(* CODESYS project ManualRequest.xml

Project tree, tasks and I/O mapping:
  visualisation ManualRequest
*)

// /ManualRequest
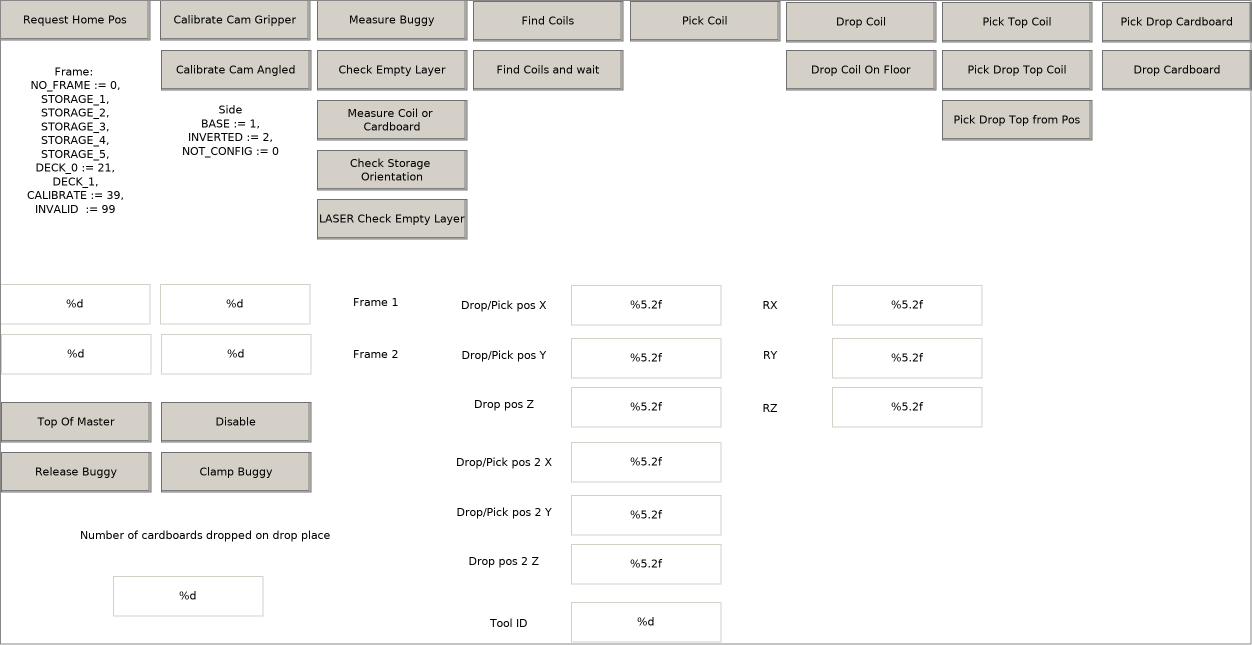
VISUALIZATION ManualRequest  // 1252x645
    Button (160,0 150x40), "Calibrate Cam Gripper", input disabled if: NOT PRG_VisuTask_10ms._fbManualCtrl.xManualMode
        tap PRG_VisuTask_10ms._fbManualCtrl._btnCalibrateCamGripper.xbtn
    Button (0,0 150x40), "Request Home Pos", input disabled if: NOT PRG_VisuTask_10ms._fbManualCtrl.xManualMode
        tap PRG_VisuTask_10ms._fbManualCtrl._btnRequestHomePos.xbtn
    Button (317,0 150x40), "Measure Buggy", input disabled if: NOT PRG_VisuTask_10ms._fbManualCtrl.xManualMode
        tap PRG_VisuTask_10ms._fbManualCtrl._btnMeasure.xbtn
    Textfield (0,284 150x40), "%d", text variable: PRG_VisuTask_10ms._fbManualCtrl._scRobotPosition.eStorage
        OnMouseUp: write the text variable via Default
    Textfield (160,284 150x40), "%d", text variable: PRG_VisuTask_10ms._fbManualCtrl._scRobotPosition.eSide
        OnMouseUp: write the text variable via Default
    Label (0,50 151x181), "Frame: NO_FRAME := 0, STORAGE_1, STORAGE_2, STORAGE_3, STORAGE_4, STORAGE_5, DECK_0 := 21, DECK_1, CALIBRATE := 39, INVALID := 99"
    Label (160,50 141x161), "Side BASE := 1, INVERTED := 2, NOT_CONFIG := 0"
    Button (473,1 150x40), "Find Coils", input disabled if: NOT PRG_VisuTask_10ms._fbManualCtrl.xManualMode
        tap PRG_VisuTask_10ms._fbManualCtrl._btnFindCoils.xbtn
    Button (630,1 150x40), "Pick Coil", input disabled if: NOT PRG_VisuTask_10ms._fbManualCtrl.xManualMode
        tap PRG_VisuTask_10ms._fbManualCtrl._btnPickCoil.xbtn
    Button (1,402 150x40), "Top Of Master", input disabled if: NOT PRG_VisuTask_10ms._fbManualCtrl.xManualMode
        tap PRG_VisuTask_10ms._fbManualCtrl._btnRequestTopOfMaster.xbtn
    Button (161,402 150x40), "Disable", input disabled if: NOT PRG_VisuTask_10ms._fbManualCtrl.xManualMode
        tap PRG_VisuTask_10ms._fbManualCtrl._btnRequestDisable.xbtn
    Button (786,2 150x40), "Drop Coil", input disabled if: NOT PRG_VisuTask_10ms._fbManualCtrl.xManualMode
        tap PRG_VisuTask_10ms._fbManualCtrl._btnDropCoil.xbtn
    Button (942,2 150x40), "Pick Top Coil", input disabled if: NOT PRG_VisuTask_10ms._fbManualCtrl.xManualMode
        tap PRG_VisuTask_10ms._fbManualCtrl._btnPickTopCoil.xbtn
    Button (1,452 150x40), "Release Buggy", input disabled if: NOT PRG_VisuTask_10ms._fbManualCtrl.xManualMode
        tap PRG_VisuTask_10ms._fbManualCtrl._btnReleaseBuggy.xbtn
    Button (161,452 150x40), "Clamp Buggy", input disabled if: NOT PRG_VisuTask_10ms._fbManualCtrl.xManualMode
        tap PRG_VisuTask_10ms._fbManualCtrl._btnClampBuggy.xbtn
    Label (445,284 118x43), "Drop/Pick pos X"
    Textfield (571,285 150x40), "%5.2f", text variable: PRG_VisuTask_10ms._fbManualCtrl._scRobotPosition.scRobotPosition.posX
        OnMouseUp: write the text variable via Default
    Textfield (571,338 150x40), "%5.2f", text variable: PRG_VisuTask_10ms._fbManualCtrl._scRobotPosition.scRobotPosition.posY
        OnMouseUp: write the text variable via Default
    Label (445,334 118x43), "Drop/Pick pos Y"
    Label (445,383 118x43), "Drop pos Z"
    Textfield (571,387 150x40), "%5.2f", text variable: PRG_VisuTask_10ms._fbManualCtrl._scRobotPosition.scRobotPosition.posZ
        OnMouseUp: write the text variable via Default
    Button (786,50 150x40), "Drop Coil On Floor", input disabled if: NOT PRG_VisuTask_10ms._fbManualCtrl.xManualMode
        tap PRG_VisuTask_10ms._fbManualCtrl._btnDropCoilOnFloor.xbtn
    Button (942,50 150x40), "Pick Drop Top Coil", input disabled if: NOT PRG_VisuTask_10ms._fbManualCtrl.xManualMode
        tap PRG_VisuTask_10ms._fbManualCtrl._btnPickDropCoil.xbtn
    Textfield (1,334 150x40), "%d", text variable: PRG_VisuTask_10ms._fbManualCtrl._scRobotPosition.eStorage2
        OnMouseUp: write the text variable via Default
    Textfield (161,334 150x40), "%d", text variable: PRG_VisuTask_10ms._fbManualCtrl._scRobotPosition.eSide2
        OnMouseUp: write the text variable via Default
    Label (317,281 118x43), "Frame 1"
    Label (317,333 118x43), "Frame 2"
    Label (445,441 118x43), "Drop/Pick pos 2 X"
    Textfield (571,442 150x40), "%5.2f", text variable: PRG_VisuTask_10ms._fbManualCtrl._scRobotPosition.scRobotPosition.pos2X
        OnMouseUp: write the text variable via Default
    Textfield (571,495 150x40), "%5.2f", text variable: PRG_VisuTask_10ms._fbManualCtrl._scRobotPosition.scRobotPosition.pos2Y
        OnMouseUp: write the text variable via Default
    Label (445,491 118x43), "Drop/Pick pos 2 Y"
    Label (445,540 118x43), "Drop pos 2 Z"
    Textfield (571,544 150x40), "%5.2f", text variable: PRG_VisuTask_10ms._fbManualCtrl._scRobotPosition.scRobotPosition.pos2Z
        OnMouseUp: write the text variable via Default
    Button (473,50 150x40), "Find Coils and wait", input disabled if: NOT PRG_VisuTask_10ms._fbManualCtrl.xManualMode
        tap PRG_VisuTask_10ms._fbManualCtrl._btnFindAndWait.xbtn
    Button (942,100 150x40), "Pick Drop Top from Pos", input disabled if: NOT PRG_VisuTask_10ms._fbManualCtrl.xManualMode
        tap PRG_VisuTask_10ms._fbManualCtrl._btnPickDropFromPos.xbtn
    Textfield (571,602 150x40), "%d", text variable: PRG_VisuTask_10ms._fbManualCtrl._scRobotPosition.scRobotPosition.ToolID
        OnMouseUp: write the text variable via Default
    Label (450,602 118x43), "Tool ID"
    Button (1102,2 150x40), "Pick Drop Cardboard", input disabled if: NOT PRG_VisuTask_10ms._fbManualCtrl.xManualMode
        tap PRG_VisuTask_10ms._fbManualCtrl._btnPickDropCardboard.xbtn
    Textfield (113,576 150x40), "%d", text variable: PersistentVars.nbrOfCardboards
        OnMouseUp: write the text variable via Default
    Label (55,502 301x67), "Number of cardboards dropped on drop place"
    Button (161,50 150x40), "Calibrate Cam Angled", input disabled if: NOT PRG_VisuTask_10ms._fbManualCtrl.xManualMode
        tap PRG_VisuTask_10ms._fbManualCtrl._btnCalibrateCamAngled.xbtn
    Button (317,50 150x40), "Check Empty Layer", input disabled if: NOT PRG_VisuTask_10ms._fbManualCtrl.xManualMode
        tap PRG_VisuTask_10ms._fbManualCtrl._btnCheckEmptyLayer.xbtn
    Button (1102,50 150x40), "Drop Cardboard", input disabled if: NOT PRG_VisuTask_10ms._fbManualCtrl.xManualMode
        tap PRG_VisuTask_10ms._fbManualCtrl._btnDropCardboard.xbtn
    Button (317,100 150x40), "Measure Coil or Cardboard", input disabled if: NOT PRG_VisuTask_10ms._fbManualCtrl.xManualMode
        tap PRG_VisuTask_10ms._fbManualCtrl._btnMeasureCoilOrCardboard.xbtn
    Label (746,284 48x43), "RX", invisible if: true
    Textfield (832,285 150x40), "%5.2f", text variable: PRG_VisuTask_10ms._fbManualCtrl._scRobotPosition.scRobotPosition.posRX, invisible if: true
        OnMouseUp: write the text variable via Default
    Textfield (832,338 150x40), "%5.2f", text variable: PRG_VisuTask_10ms._fbManualCtrl._scRobotPosition.scRobotPosition.posRY, invisible if: true
        OnMouseUp: write the text variable via Default
    Textfield (832,387 150x40), "%5.2f", text variable: PRG_VisuTask_10ms._fbManualCtrl._scRobotPosition.scRobotPosition.posRZ, invisible if: true
        OnMouseUp: write the text variable via Default
    Label (746,334 48x43), "RY", invisible if: true
    Label (746,387 48x43), "RZ", invisible if: true
    Button (317,150 150x40), "Check Storage Orientation", input disabled if: NOT PRG_VisuTask_10ms._fbManualCtrl.xManualMode
        tap PRG_VisuTask_10ms._fbManualCtrl._btnCheckStorageOrientation.xbtn
    Button (317,199 150x40), "LASER Check Empty Layer", input disabled if: NOT PRG_VisuTask_10ms._fbManualCtrl.xManualMode
        tap PRG_VisuTask_10ms._fbManualCtrl._btnCheckEmptyLayerLaser.xbtn
END_VISUALIZATION
